// TIA Portal V21 export
DATA_BLOCK "HMI_Steuerung_DB"   // DB10
{ S7_Optimized_Access := 'TRUE' }
// stored: MemoryReserve 100
   VAR
      Pos_v : LReal;
      Vel_v : LReal;
      Vel_absolut_v : LReal;   // angepasste Geschwindigkeit für vertikale Achse in %
      Pos_h : LReal;
      Vel_h : LReal;
      Vel_absolut_h : LReal;   // angepasste Geschwindigkeit für horizontale Achse in %
      Pos_z : LReal;
      Vel_z : LReal;
      jog_mode_hoch : Bool;
      jog_mode_runter : Bool;
      jog_mode_rechts : Bool;
      jog_mode_links : Bool;
      EnableSwitch : Bool;
      ExecuteMode : Bool;
      StopMode : Bool;
      Inkrement_relativ : LReal;
      relativ_hoch : Bool;
      relativ_runter : Bool;
      relativ_rechts : Bool;
      relativ_links : Bool;
      Set_Ventil_A : Bool;
   END_VAR
BEGIN
END_DATA_BLOCK
